ABB RAPID module: ProbeProg.mod

%%%
  VERSION:1
  LANGUAGE:ENGLISH
%%%
MODULE MOD_ProbeProg

    ! -------------------------------
    ! Define customized variables here
    ! ...

	! Tool variables:
	PERS tooldata ProbeTool := [TRUE,[[0.000,0.000,100.000],[1.00000000,0.00000000,0.00000000,0.00000000]],[1,[0,0,20],[1,0,0,0],0,0,0.005]];

	! Reference variables:
	PERS wobjdata ProbeFrameRenamed := [FALSE, TRUE, "", [[0,0,0],[1,0,0,0]],[[100.000,-1000.000,300.000],[0.70710678,0.00000000,0.00000000,0.70710678]]];

	PROC Main()
		ConfJ \On;
		ConfL \Off;
		! Program generated by RoboCraft v1.0 for ABB IRB 120-3/0.6 on XX/XX/XXXX 14:46:38
		! Using nominal kinematics.
		MoveAbsJ [[0.000000,-10.000000,20.000000,0.000000,30.000000,0.000000],[9E+09,9E+09,9E+09,9E+09,9E+09,9E+09]],[250.00,500,5000,1000],z5,ProbeTool \WObj:=ProbeFrameRenamed;
		MoveL [[1050.000,-294.442,161.833],[0.29883624,0.64085638,0.64085638,-0.29883624],[0,0,0,0],[9E+09,9E+09,9E+09,9E+09,9E+09,9E+09]],[250.00,500,5000,1000],z5,ProbeTool \WObj:=ProbeFrameRenamed;
		MoveAbsJ [[20.000000,-10.000000,20.000000,0.000000,30.000000,0.000000],[9E+09,9E+09,9E+09,9E+09,9E+09,9E+09]],[250.00,500,5000,1000],z5,ProbeTool \WObj:=ProbeFrameRenamed;
		WaitTime 0.500;
		TPWrite "Hello from probe";
		! a comment
		SetDO D_OUT_1, 1;
		WaitDI D_IN_2, 1, \MaxTime:=1.0;
		SubProgram;
	ENDPROC

ENDMODULE
